SUBAPPLICATION IN_UP (* Subapplication Type *)
  (* Standard: 61499-2 *)
  (* Version 1.0, 2023-02-06, franz *)
  IMPORT BlinkMarine::io::DI::PKP_2200_LI_DI::Invalid;
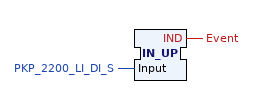
  EVENT_OUTPUT
    IND;
  END_EVENT
  VAR_INPUT
    Input : BlinkMarine::io::DI::PKP_2200_LI_DI_S := Invalid;
  END_VAR
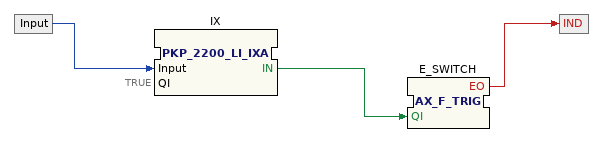
  FBS
    E_SWITCH : adapter::events::unidirectional::AX_F_TRIG;
    IX : BlinkMarine::io::DI::PKP_2200_LI_IXA(QI := TRUE);
  END_FBS
  EVENT_CONNECTIONS
    E_SWITCH.EO TO IND;
  END_CONNECTIONS
  DATA_CONNECTIONS
    Input TO IX.Input;
  END_CONNECTIONS
  ADAPTER_CONNECTIONS
    IX.IN TO E_SWITCH.QI;
  END_CONNECTIONS
END_SUBAPPLICATION
